(* IEC 61131-3 sources: openplc-editor-canopen/e2e/fixtures/canopen-generic-io/project/pous/programs, 1 file *)

(* ---- main.st ---- *)
PROGRAM main
  VAR
    in0 AT %IX0.0 : BOOL;
    in1 AT %IX0.1 : BOOL;
    in2 AT %IX0.2 : BOOL;
    in3 AT %IX0.3 : BOOL;
    in4 AT %IX0.4 : BOOL;
    in5 AT %IX0.5 : BOOL;
    in6 AT %IX0.6 : BOOL;
    in7 AT %IX0.7 : BOOL;
    out0 AT %QX0.0 : BOOL;
    out1 AT %QX0.1 : BOOL;
    out2 AT %QX0.2 : BOOL;
    out3 AT %QX0.3 : BOOL;
    out4 AT %QX0.4 : BOOL;
    out5 AT %QX0.5 : BOOL;
    out6 AT %QX0.6 : BOOL;
    out7 AT %QX0.7 : BOOL;
  END_VAR

out0 := in0;
out1 := in1;
out2 := in2;
out3 := in3;
out4 := in4;
out5 := in5;
out6 := in6;
out7 := in7;

END_PROGRAM
